Universal Robots URScript: PgProg.script

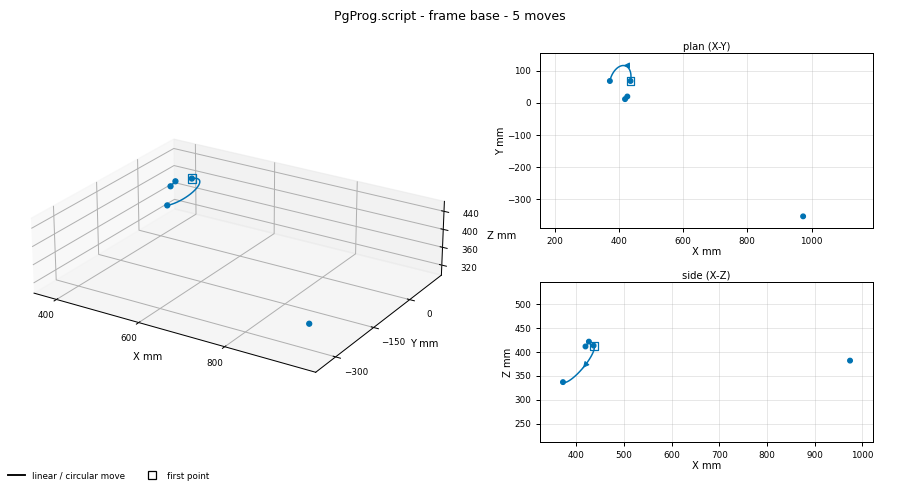
[picture p0: tool path of PgProg.script in frame base, 5 of 9 moves have a stored position in this frame; points joined in program order, loops and branches not executed]
def PgProg():
  # Global parameters:
  global speed_ms    = 0.250
  global speed_rads  = 0.750
  global accel_mss   = 1.200
  global accel_radss = 1.200
  global blend_radius_m = 0.001
  global ref_frame = p[0,0,0,0,0,0]

  #
  # TO REMOVE HEADER:
  # Go to "Program" -> "Post-Processor Editor"
  # Select "Universal Robots"
  # Set "INCLUDE_HEADER" to "False"
  #
  #--------------------------
  # Add any default subprograms here
  # For example, to drive a gripper as a program call:
  # def Gripper_Open():
  #   ...
  # end
  #
  # Example to drive a spray gun:
  def SprayOn(value):
    # use the value as an output:
    DO_SPRAY = 5
    if value == 0:
      set_standard_digital_out(DO_SPRAY, False)
    else:
      set_standard_digital_out(DO_SPRAY, True)
    end
  end

  # Example to drive an extruder:
  def Extruder(value):
    # use the value as an output:
    if value < 0:
      # stop extruder
    else:
      # start extruder
    end
  end

  # Example to move an external axis
  def MoveAxis(value):
    # use the value as an output:
    DO_AXIS_1 = 1
    DI_AXIS_1 = 1
    if value <= 0:
      set_standard_digital_out(DO_AXIS_1, False)

      # Wait for digital input to change state
      #while (get_standard_digital_in(DI_AXIS_1) != False):
      #  sync()
      #end
    else:
      set_standard_digital_out(DO_AXIS_1, True)

      # Wait for digital input to change state
      #while (get_standard_digital_in(DI_AXIS_1) != True):
      #  sync()
      #end
    end
  end
  #--------------------------


  # Main program:
  # Program generated by RoboDK v6.0.7 for UR10 on XX/XX/XXXX 18:00:00
  # Using nominal kinematics.
  ref_frame = p[1.234570, -0.098765, 0.050500, 0.000000, 0.000000, 0.523599]
  set_tcp(p[0.010000, 0.020000, 0.150000, 0.261799, 0.000000, 0.000000])
  blend_radius_m = 0.005
  movej([0.000000, -0.174533, 0.349066, 0.000000, 0.523599, 0.000000],accel_radss,speed_rads,t=0,r=0)
  movel(pose_trans(ref_frame,p[-0.607850, 0.543849, 0.363215, 0.731956, 2.185937, -0.570291]),accel_mss,speed_ms,t=0,r=0.005)
  movec(pose_trans(ref_frame,p[-0.602951, 0.596788, 0.316595, 0.731956, 2.185937, -0.570291]),pose_trans(ref_frame,p[-0.663517, 0.575988, 0.286611, 0.731956, 2.185937, -0.570291]),accel_mss,speed_ms,r=0.005)
  movej([0.349066, -0.174533, 0.349066, 0.000000, 0.523599, 0.000000],accel_radss,speed_rads,t=0,r=0)
  accel_radss = 2.094
  speed_rads  = 1.047
  accel_mss   = 0.800
  speed_ms    = 0.100
  movel(pose_trans(ref_frame,p[-0.650861, 0.503437, 0.361399, 0.731956, 2.185937, -0.570291]),accel_mss,speed_ms,t=0,r=0)
  blend_radius_m = 0.000
  movel(pose_trans(ref_frame,p[-0.640584, 0.506980, 0.371534, 0.731956, 2.185937, -0.570291]),accel_mss,speed_ms,t=0,r=0.000)
  sleep(0.500)
  halt() # reimplement this function to force stop
  popup("Hello from postgen","Message",False,False,blocking=True)
  # a comment
  SubProgram()
  CustomCode(42)
  ThreadProg
  set_standard_digital_out(1, True)
  Valve = 0
  set_standard_analog_out(3, 2.5)
  while (get_standard_digital_in(2) != True):
    sync()
  end
  while (get_standard_digital_in(4) != False):
    sync()
  end
  set_tcp(p[0.000000, 0.000000, 0.200000, 0.000000, 0.000000, 0.000000])
  movej([0.000000, -0.174533, 0.349066, 0.000000, 0.523599, 0.000000],accel_radss,speed_rads,t=0,r=0.000)
  movej([0.174533, -0.087266, 0.436332, 0.087266, 0.610865, 0.087266],accel_radss,speed_rads,t=0,r=0)
  movel(pose_trans(ref_frame,p[-0.353026, -0.090135, 0.331702, 0.124818, 2.423541, -0.239517]),accel_mss,speed_ms,t=0,r=0)
  # End of main program
end

PgProg()
